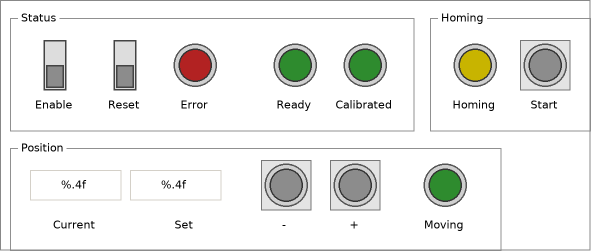
VISUALIZATION Focus  // 591x251
    GroupBox (10,10 404x121), "Status"
        DipSwitch (20,30 50x50), variable: MAIN.focusControl.bEnable, behaviour: TOGGLE, style: Switch-DipSwitch-Gray
        DipSwitch (90,30 50x50), variable: MAIN.focusControl.bReset, behaviour: TOGGLE, style: Switch-DipSwitch-Gray
        Lamp1 (160,30 50x50), variable: MAIN.focusControl.bError, style: Lamp-Lamp1-Red
        Lamp1 (260,30 50x50), variable: MAIN.focusControl.bReady, style: Lamp-Lamp1-Green
        Lamp1 (330,30 50x50), variable: MAIN.focusControl.bCalibrated, style: Lamp-Lamp1-Green
        Label (10,80 68x30), "Enable"
        Label (80,80 68x30), "Reset"
        Label (150,80 68x30), "Error"
        Label (250,80 68x30), "Ready"
        Label (320,80 68x30), "Calibrated"
    GroupBox (430,10 161x121), "Homing"
        Lamp1 (20,30 50x50), variable: MAIN.focusControl.bHomeAxis, style: Lamp-Lamp1-Yellow
        Label (10,80 68x30), "Homing"
        PushSwitch (90,30 50x50), variable: MAIN.focusControl.bHomeAxis, behaviour: TOGGLE, style: Switch-PushSwitch-Gray
        Label (80,80 68x30), "Start"
    GroupBox (10,140 491x111), "Position"
        Textfield (20,30 91x30), "%.4f", text variable: MAIN.focusControl.fActualPosition
        Label (30,70 68x30), "Current"
        Textfield (120,30 91x30), "%.4f", text variable: MAIN.focusControl.fPosition
            OnMouseUp: write the text variable via InputWithLimits, min MAIN.focusControl.fMinPosition, max MAIN.focusControl.fMaxPosition
        PushSwitch (251,20 50x50), variable: MAIN.focusControl.bMoveNeg, behaviour: TOGGLE, style: Switch-PushSwitch-Gray
        PushSwitch (320,20 50x50), variable: MAIN.focusControl.bMovePos, behaviour: TOGGLE, style: Switch-PushSwitch-Gray
        Label (240,70 68x30), "-"
        Label (310,70 68x30), "+"
        Label (140,70 68x30), "Set"
        Lamp1 (410,20 50x50), variable: MAIN.focusControl.bMoveAxis, style: Lamp-Lamp1-Green
        Label (400,70 68x30), "Moving"
END_VISUALIZATION

(* stored: Version 1.1.0.1, ProductVersion 3.1.4024.15
   Visu Focus: Id {61a00a5d-5dbf-408f-af24-517c83e1ab5f} *)
